Staubli VAL3: resetMoveId.pgx

public program resetMoveId()
  local num l_nNextId
begin
  //reset move id to avoid move id overflow
  l_nNextId=nextMoveId()
  if l_nNextId>=nMoveIdMax
    setMoveId(0)
  endIf
end
